(* IEC 61131-3 sources: plcfuzz/testcases/matiec/experimental, 3 files *)

(* ---- function_block_method.st ---- *)
FUNCTION_BLOCK Accumulator
  VAR
    Total : INT := 0;
  END_VAR

  Total := Total;

  METHOD PUBLIC Add : INT
    VAR_INPUT
      Delta : INT;
    END_VAR
    Total := Total + Delta;
    Add := Total;
  END_METHOD
END_FUNCTION_BLOCK

PROGRAM MethodDemo
  VAR
    Instance : Accumulator;
    Result : INT;
  END_VAR

  Result := Instance.Add(Delta := 2);
END_PROGRAM

CONFIGURATION Config0
  RESOURCE Res0 ON PLC
    TASK MainTask(INTERVAL := T#100ms, PRIORITY := 0);
    PROGRAM Instance0 WITH MainTask : MethodDemo;
  END_RESOURCE
END_CONFIGURATION

(* ---- utf8_string.st ---- *)
PROGRAM Utf8Status
  VAR
    StatusMessage : STRING := '设备就绪🚀';
  END_VAR

  StatusMessage := StatusMessage;
END_PROGRAM

CONFIGURATION Config0
  RESOURCE Res0 ON PLC
    TASK MainTask(INTERVAL := T#100ms, PRIORITY := 0);
    PROGRAM Instance0 WITH MainTask : Utf8Status;
  END_RESOURCE
END_CONFIGURATION

(* ---- variable_access.st ---- *)
PROGRAM AccessDemo
  VAR_OUTPUT
    CurrentValue : INT;
  END_VAR
  CurrentValue := CurrentValue + 1;
END_PROGRAM

CONFIGURATION AccessConfig
  VAR_GLOBAL
    Setpoint : INT := 100;
  END_VAR

  RESOURCE Res0 ON PLC
    TASK MainTask(INTERVAL := T#100ms, PRIORITY := 0);
    PROGRAM Instance0 WITH MainTask : AccessDemo;
  END_RESOURCE

  VAR_ACCESS
    RemoteSetpoint : Setpoint : INT READ_WRITE;
    MonitorValue : Res0.Instance0.CurrentValue : INT READ_ONLY;
  END_VAR
END_CONFIGURATION
